DATA_BLOCK "FRK_ClassScratch"
{ S7_Optimized_Access := 'TRUE' }
VERSION : 0.1
NON_RETAIN
VAR
    Blank {ExternalAccessible := 'False'; ExternalVisible := 'False'; ExternalWritable := 'False'} : "ST_DataClassPolicy";
END_VAR
BEGIN
END_DATA_BLOCK
